Fanuc KAREL source: kt00549.KL

-- PROVISIONAL review KL for V1013-1; original PC SHA256 6eb2e87c121ca0f93095d2ff827b446e0882d53215651c1cf600617c01898fa6
-- Incomplete behavior may be omitted. Consult companion uncertainty JSON. Do not deploy.
PROGRAM KT00549
%NOLOCKGROUP
-- UNRESOLVED_DECL P1 type=000199
-- UNRESOLVED_DECL P2 type=000199
-- UNRESOLVED_DECL OUT type=000101
BEGIN
  -- UNRESOLVED_PC offsets 5-39; opcodes 49,7E,49,7E,60,4A
  -- UNRESOLVED_PC offsets 44-48; opcodes 7F
END KT00549
